// TIA Portal V19 export
TYPE "PidL.HMI"
   STRUCT
      identName : String;
      comment : String;
      AutModOp : Bool;
      ManModOp : Bool;
      LocModOp : Bool;
      OosModOp : Bool;
      ResetOp : Bool;
      MonitorOn : Bool;
      ExtModOp : Bool;
      IntModOp : Bool;
      SpInt : Real;
      Man : Real;
      PermissionLog { S7_SetPoint := 'True'} : "PidL.Permission";
      Status { S7_SetPoint := 'True'} : "PidL.Status";
      PIDConfig { S7_SetPoint := 'True'} : "PidL.PIDConfig";
      Alarms { S7_SetPoint := 'True'} : "AnaMon.HMI";
   END_STRUCT;
END_TYPE
